Fanuc KAREL source: KB00054.KL

PROGRAM KB00054
%NOLOCKGROUP
VAR
  P1: INTEGER
  P2: INTEGER
  P3: INTEGER
BEGIN
  P1 = 1
  P2 = 1
  P3 = 1
  DAQ_CHECKP(P1, P2, P3)
END KB00054
